PROGRAM main
  VAR
    SCADA_ALARM_ACTIVATE AT %QX0.0 : BOOL;
    PUB_REMOTE_ONLY AT %QX0.1 : BOOL;
    PUB_MANUAL_PULL_TRIGGERED AT %QX0.2 : BOOL;
    PUB_FLAME_DETECTED AT %QX0.3 : BOOL;
    PUB_GAS_SMOKE_ALERT AT %QX0.4 : BOOL;
    PUB_GAS_RAW_VALUE AT %QW0 : UINT;
    PUB_HEARTBEAT AT %QW1 : UINT;
    PUB_RECONNECT_COUNT AT %QW2 : UINT;
    ALARM_ACTIVATE AT %QX100.0 : BOOL;
    MANUAL_PULL_TRIGGERED AT %IX100.0 : BOOL;
    FLAME_DETECTED AT %IX100.1 : BOOL;
    GAS_SMOKE_ALERT AT %IX100.2 : BOOL;
    GAS_RAW_VALUE AT %IW100 : UINT;
    HEARTBEAT AT %IW101 : UINT;
    RECONNECT_COUNT AT %IW102 : UINT;
  END_VAR

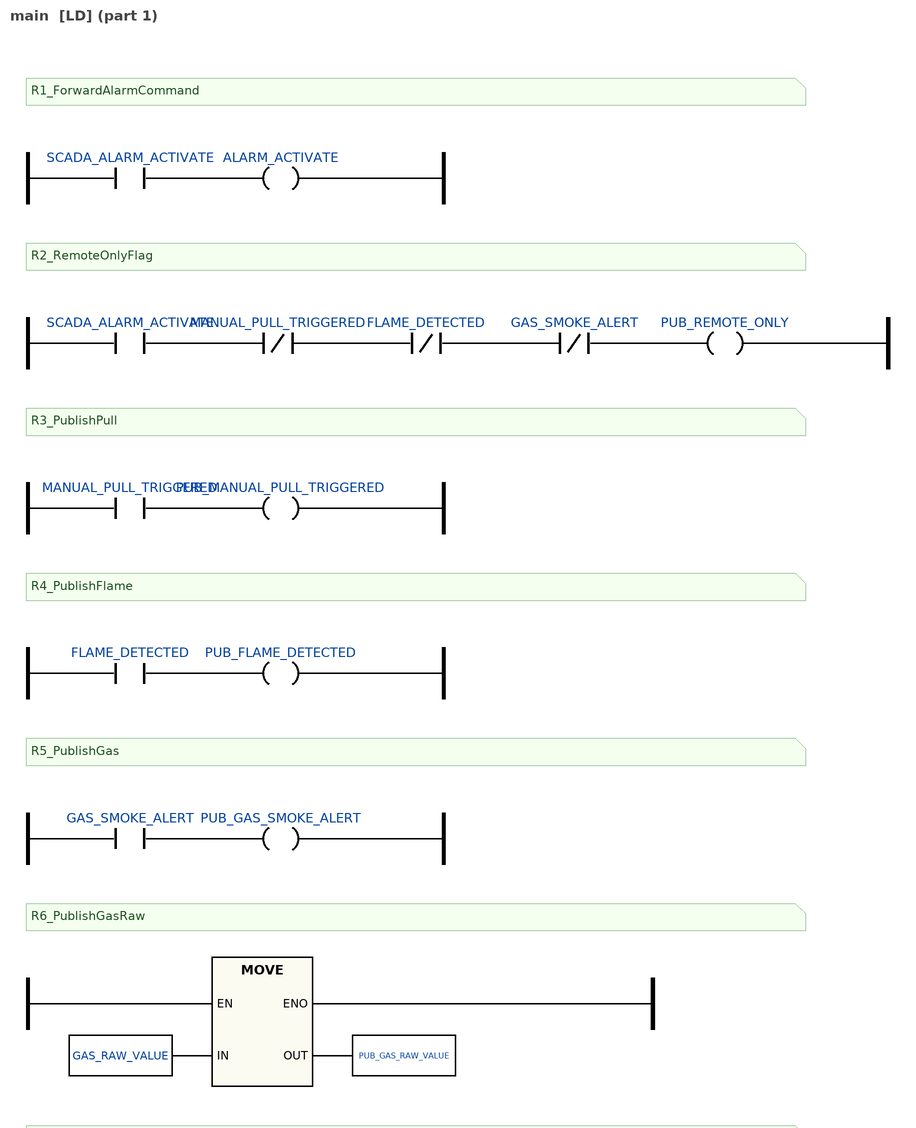
(* LD diagram, written out as Structured Text *)
(* R1_ForwardAlarmCommand *)
ALARM_ACTIVATE := SCADA_ALARM_ACTIVATE;
(* R2_RemoteOnlyFlag *)
PUB_REMOTE_ONLY := SCADA_ALARM_ACTIVATE AND NOT MANUAL_PULL_TRIGGERED AND NOT FLAME_DETECTED AND NOT GAS_SMOKE_ALERT;
(* R3_PublishPull *)
PUB_MANUAL_PULL_TRIGGERED := MANUAL_PULL_TRIGGERED;
(* R4_PublishFlame *)
PUB_FLAME_DETECTED := FLAME_DETECTED;
(* R5_PublishGas *)
PUB_GAS_SMOKE_ALERT := GAS_SMOKE_ALERT;
(* R6_PublishGasRaw *)
PUB_GAS_RAW_VALUE := GAS_RAW_VALUE;
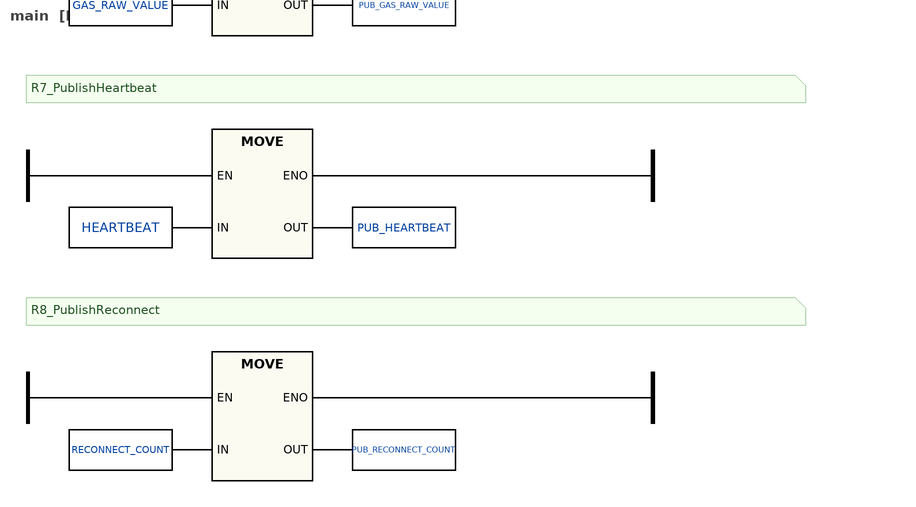
(* R7_PublishHeartbeat *)
PUB_HEARTBEAT := HEARTBEAT;
(* R8_PublishReconnect *)
PUB_RECONNECT_COUNT := RECONNECT_COUNT;
END_PROGRAM
